(* CODESYS project BODAS-RC18-12_27-18_40-DSA.library
   Company: Bosch Rexroth AG
   DefaultNamespace: BODAS-API-RC18-12_27-18_40-DSA
   Version: 2.3.0
   DocFormat: reStructuredText
   Description: User library to use BODAS-BDL services (API) for RC40.
   Title: BODAS_RC18-12_27-18_40-DSA

Project tree, tasks and I/O mapping:
  DSA/
    API/
      function bds_snsrDsa_getTemp [ST]
      function bds_snsrDsa_cfgSpdAndDir [ST]
      function bds_snsrDsa_getSpdAndDir [ST]
    ENUM/
      data type bds_snsrDsa_status_te
      data type bds_snsrDsa_dir_te
    STRUCT/
      data type bds_snsrDsa_cfgSpdAndDir_ts
      data type bds_snsrDsa_statusDiag_tb
      data type bds_snsrDsa_getSpdAndDir_ts
      data type bds_snsrDsa_getTemp_ts
*)

// DSA/ENUM/bds_snsrDsa_status_te
{attribute 'external_name' := 'cmp_rts_bds_snsrDsa_status_te'}
TYPE bds_snsrDsa_status_te : 
(
    bds_snsrDsa_ok_E := 0,                (* API function call is ok *)
    bds_snsrDsa_outOfRange_E := 1,        (* The detected frequency for CW, CCW or calculated rpm are out of range *)
    bds_snsrDsa_frzn_E := 2,              (* Provided rpm value is frozen *)
    bds_snsrDsa_standStill_E := 3,        (* Detected rpm value is 0 and freezetime is elapsed *)
    bds_snsrDsa_err_E := 4,               (* Diagnostic error (SCG, SCB, OL detected or hardware error) *)
    bds_snsrDsa_invldConfig_E := 5,       (* Invalid configuration like no. of teeth is out of range *)
    bds_snsrDsa_notConfig_E := 6,         (* Not configured e.g. resistance input is not configured *)
    bds_snsrDsa_invldPrm_E := 7           (* Wrong parameter e.g. DSA instance is not configured *)
) USINT;
END_TYPE

// DSA/STRUCT/bds_snsrDsa_cfgSpdAndDir_ts
{attribute 'external_name' := 'cmp_rts_bds_snsrDsa_cfgSpdAndDir_ts'}
TYPE bds_snsrDsa_cfgSpdAndDir_ts : STRUCT
    stsApi_e : bds_snsrDsa_status_te;           (* Return status of Api call *)
END_STRUCT
END_TYPE

// DSA/STRUCT/bds_snsrDsa_statusDiag_tb
{attribute 'external_name' := 'cmp_rts_bds_snsrDsa_statusDiag_tb'}
{attribute 'size' := '32'}
TYPE bds_snsrDsa_statusDiag_tb : STRUCT
    stErrSCB_b1 : BIT;     (* Status of short cut to battery *)
    stErrSCG_b1 : BIT;     (* Status of short cut to ground *)
    stErrOL_b1 : BIT;      (* Status of open load *)
    stErrOT_b1 : BIT;      (* Status of over temperature *)
    stErrUT_b1 : BIT;      (* Status of under temperature *)
    stErrHw_b1 : BIT;      (* Status of hardware error *)
	resd1_b : ARRAY[0..2] OF BYTE;      (* Reserved *)
END_STRUCT
END_TYPE

// DSA/ENUM/bds_snsrDsa_dir_te
{attribute 'external_name' := 'cmp_rts_bds_snsrDsa_dir_te'}
TYPE bds_snsrDsa_dir_te : 
(
    bds_snsrDsa_dirUnkown_E := 0,           (* Rotation direction is not known *)
    bds_snsrDsa_dirClockwise_E := 1,        (* Rotation direction is clockwise *)
    bds_snsrDsa_dirCounterClockwise_E := 2, (* Rotation direction is counter-clockwise *)
    bds_snsrDsa_dirImpsChgErr_E := 3        (* Rotation direction is implausible *)
) USINT;
END_TYPE

// DSA/STRUCT/bds_snsrDsa_getSpdAndDir_ts
{attribute 'external_name' := 'cmp_rts_bds_snsrDsa_getSpdAndDir_ts'}
TYPE bds_snsrDsa_getSpdAndDir_ts : STRUCT
    statusDiag_b : bds_snsrDsa_statusDiag_tb;   (* Diagnostic information of sensor *)
    spd_dRpm_u32 : UDINT;                       (* Rotation speed in deci Rpm *)
    dir_e : bds_snsrDsa_dir_te;                 (* Rotation direction of sensor *)
    stsApi_e : bds_snsrDsa_status_te;           (* Return status of API call *)
END_STRUCT
END_TYPE

// DSA/STRUCT/bds_snsrDsa_getTemp_ts
{attribute 'external_name' := 'cmp_rts_bds_snsrDsa_getTemp_ts'}
TYPE bds_snsrDsa_getTemp_ts : STRUCT
    stsApi_e : bds_snsrDsa_status_te;           (* Return status of Api call *)
    statusDiag_b : bds_snsrDsa_statusDiag_tb;   (* Diagnostic information of temperature *)
    temp_degC_s32 : DINT;                       (* Temperature in degrees Celsius *)
END_STRUCT
END_TYPE

// DSA/API/bds_snsrDsa_getTemp
/// The bds_snsrDsa_getTemp API function provides temperature in degree celsius and diagnostic status of a particular DSA sensor instance.
///
///  
///==================================================================		  			===================================================================================================
///Return value    								  									     Description
///==================================================================		  			===================================================================================================
/// bds_snsrDsa_getTemp_ts																 The return structure containing the status of API function call, temperature in degree celsius and diagnostic information of a particular DSA sensor instance. For detailed information, please refer to chapter 																
///
///==================================================================		   			===================================================================================================
///
///=======
///Code Example:
///=======
///============================================================================
///
/// PROGRAM OsInitProc
///VAR
///
///    bds_snsrDsa_getTemp_s : bds_snsrDsa_getTemp_ts;
///	
///    bds_snsrDsa_inst_e : bds_snsrDsa_inst_te;
///	
///    temp_degC_s32 : DINT;
///	
///END_VAR
///
///bds_snsrDsa_inst_e := bds_snsrDsa_inst_te.DrvPumpSpeed_E;
///
///bds_snsrDsa_getTemp_s := bds_snsrDsa_getTemp(bds_snsrDsa_inst_e);
///
///IF bds_snsrDsa_ok_E = bds_snsrDsa_getTemp_s.statusApi_e THEN
///
///    (* save the actual temperature in degree celsius *)
///	
///    temp_degC_s32 := bds_snsrDsa_getTemp_s.temp_degC_s32;
///	
///ELSE
///
///    (* error handling *)
///	
///END_IF;
/// END_PROGRAM
///
///
///============================================================================
{attribute 'external_name' := 'cmp_rts_bds_snsrDsa_getTemp'}
FUNCTION bds_snsrDsa_getTemp : bds_snsrDsa_getTemp_ts
VAR_INPUT
///The DSA sensor instance name.
snsrDsaInst_e: USINT;
END_VAR

END_FUNCTION

// DSA/API/bds_snsrDsa_cfgSpdAndDir
/// The bds_snsrDsa_cfgSpdAndDir API function configures the number of encoder wheel teeth.
///
///==================================================================		  			===================================================================================================
///Return value    								  									     Description
///==================================================================		  			===================================================================================================
/// bds_snsrDsa_cfgSpdAndDir_ts															 The return structure containing the status of API function call.																
///
///==================================================================		   			===================================================================================================
///
///=======
///Code Example:
///=======
///============================================================================
///
///PROGRAM OsInitProc
///VAR
///
///    bds_snsrDsa_cfgSpdAndDir_s : bds_snsrDsa_cfgSpdAndDir_ts;
///	
///    bds_snsrDsa_inst_e : bds_snsrDsa_inst_te;
///	
///    nrOfTeeth_u16 : UINT := 75;
///	
///END_VAR
///
/// bds_snsrDsa_inst_e := bds_snsrDsa_inst_te.DrvPumpSpeed_E;
///
/// bds_snsrDsa_cfgSpdAndDir_s := bds_snsrDsa_cfgSpdAndDir(bds_snsrDsa_inst_e, nrOfTeeth_u16);
///
///IF bds_snsrDsa_ok_E = bds_snsrDsa_cfgSpdAndDir_s.statusApi_e THEN
///
///    (* configuration of DST sensor instance is successful *)
///	
///ELSE
///
///    (* error handling *)
///	
///END_IF;
/// END_PROGRAM
///
///============================================================================

{attribute 'external_name' := 'cmp_rts_bds_snsrDsa_cfgSpdAndDir'}
FUNCTION bds_snsrDsa_cfgSpdAndDir : bds_snsrDsa_cfgSpdAndDir_ts
VAR_INPUT
///The DSA sensor instance name.
snsrDsaInst_e: USINT;
///The number of wheel teeth for a particular DSA sensor instance.
///The range of wheel teeth is from 0 to 1000.
nrOfTeeth_u16: UINT;
END_VAR

END_FUNCTION

// DSA/API/bds_snsrDsa_getSpdAndDir
/// The bds_snsrDsa_getSpdAndDir API function provides calculated rotation speed with resolution of 0.1 rpm, rotation direction and diagnostic status of a particular DSA sensor instance.
///
///Remarks
///
/// A configuration function bds_snsrDsa_cfgSpdAndDir is necessary, because calculation of rotation speed is based on number of wheel teeth.
///
///  
///==================================================================		  			===================================================================================================
///Return value    								  									     Description
///==================================================================		  			===================================================================================================
/// bds_snsrDsa_getSpdAndDir_ts															  containing the status of API function call, wheel rotation speed in deci-rpm, wheel rotation direction and diagnostic information of a particular DSA sensor instance. For detailed information, please refer to chapter DSA.																
///
///==================================================================		   			===================================================================================================
///
///=======
///Code Example:
///=======
///============================================================================
///
/// PROGRAM OsInitProc
///VAR
///
///    bds_snsrDsa_getSpdAndDir_s : bds_snsrDsa_getSpdAndDir_ts;
///	
///    bds_snsrDsa_inst_e : bds_snsrDsa_inst_te;
///	
///    spd_dRpm_u32 : UDINT;
///	
///    rotDir_u8 : bds_snsrDsa_dir_te;
///	
///END_VAR
///
///bds_snsrDsa_inst_e := bds_snsrDsa_inst_te.DrvPumpSpeed_E;
///
///bds_snsrDsa_getSpdAndDir_s := bds_snsrDsa_getSpdAndDir(bds_snsrDsa_inst_e);
///
///IF bds_snsrDst_ok_E = bds_snsrDsa_getSpdAndDir_s.statusApi_e THEN
///
///    (* save the actual wheel speed and rotation direction *)
///	
///    spd_dRpm_u32 := bds_snsrDsa_getSpdAndDir_s.spd_dRpm_u32;
///	
///    rotDir_u8 := bds_snsrDsa_getSpdAndDir_s.dir_e;
///	
///ELSE
///
///    (* error handling *)
///	
///END_IF;
/// END_PROGRAM
///
///
///============================================================================
{attribute 'external_name' := 'cmp_rts_bds_snsrDsa_getSpdAndDir'}
FUNCTION bds_snsrDsa_getSpdAndDir : bds_snsrDsa_getSpdAndDir_ts
VAR_INPUT
///The DSA sensor instance name.
snsrDsaInst_e: USINT;
END_VAR

END_FUNCTION
